TYPE ST_DeviceId :
STRUCT
    sId      : UINT;
    sName    : STRING(32);
    sRoom    : STRING(32);
    bEnabled : BOOL := TRUE;
END_STRUCT
END_TYPE

(* stored: Version 1.1.0.1, ProductVersion 3.1.4026.20
   DUT ST_DeviceId: Id {44444444-4444-4444-8444-444444444444} *)
